(* PLC project GeneratedProgram, SafePLC-Gen SafePLC-Gen Multimodal 1.0 *)
(* stored: creationDateTime 2026-04-25T11:55:04.001507Z *)

PROGRAM GeneratedProgram
  VAR
    FirstScan : BOOL;
    TICSA_4750_03_Scaled : REAL;
    PICSA_4712_02_Scaled : REAL;
    PI_4712_01_Scaled : REAL;
    TICSA_4750_03_EU_Min : REAL;
    TICSA_4750_03_EU_Span : REAL;
    PICSA_4712_02_EU_Min : REAL;
    PICSA_4712_02_EU_Span : REAL;
    PI_4712_01_EU_Min : REAL;
    PI_4712_01_EU_Span : REAL;
    TICSA_4750_03_HH_SP : REAL;
    TICSA_4750_03_H_SP : REAL;
    TICSA_4750_03_L_SP : REAL;
    TICSA_4750_03_LL_SP : REAL;
    TICSA_4750_03_Deadband : REAL;
    PICSA_4712_02_HH_SP : REAL;
    PICSA_4712_02_H_SP : REAL;
    PICSA_4712_02_L_SP : REAL;
    PICSA_4712_02_LL_SP : REAL;
    PICSA_4712_02_Deadband : REAL;
    PI_4712_01_HH_SP : REAL;
    PI_4712_01_H_SP : REAL;
    PI_4712_01_L_SP : REAL;
    PI_4712_01_LL_SP : REAL;
    PI_4712_01_Deadband : REAL;
    TICSA_4750_03_HH_Ack : BOOL;
    TICSA_4750_03_LL_Ack : BOOL;
    PICSA_4712_02_HH_Ack : BOOL;
    PICSA_4712_02_LL_Ack : BOOL;
    PI_4712_01_HH_Ack : BOOL;
    PI_4712_01_LL_Ack : BOOL;
    TICSA_4750_03_LL_Latched : BOOL;
    PICSA_4712_02_HH_Latched : BOOL;
    PICSA_4712_02_LL_Latched : BOOL;
    PI_4712_01_HH_Latched : BOOL;
    PI_4712_01_LL_Latched : BOOL;
    TICSA_4750_03_HH : BOOL;
    TICSA_4750_03_LL : BOOL;
    TICSA_4750_03_H : BOOL;
    TICSA_4750_03_L : BOOL;
    PICSA_4712_02_HH : BOOL;
    PICSA_4712_02_LL : BOOL;
    PICSA_4712_02_H : BOOL;
    PICSA_4712_02_L : BOOL;
    PI_4712_01_HH : BOOL;
    PI_4712_01_LL : BOOL;
    PI_4712_01_H : BOOL;
    PI_4712_01_L : BOOL;
    LOOP_4750_03_TRIP : BOOL;
    LOOP_4712_02_TRIP : BOOL;
    LOOP_104_01_TRIP : BOOL;
    SV_104_01_HH : BOOL;
    SV_104_01_LL : BOOL;
    SAFE_STATE : BOOL;
    TIC_SP : REAL;
    TIC_Error : REAL;
    TIC_Integral : REAL;
    TIC_Kp : REAL;
    TIC_Ki : REAL;
    TIC_Output : REAL;
    PIC_SP : REAL;
    PIC_Error : REAL;
    PIC_Integral : REAL;
    PIC_Kp : REAL;
    PIC_Ki : REAL;
    PIC_Output : REAL;
    HV_MNb_47121 : BOOL;
    HV_MNb_47122 : BOOL;
    HV_75SA21 : BOOL;
    CV_73KH12_50_inlet : BOOL;
    HV_MNc_47125_block : BOOL;
    HV_MNc_47126 : BOOL;
    HV_73KH12_50_main : BOOL;
    HV_QSa_47140 : BOOL;
    HV_QSb_47141 : BOOL;
    HV_MNc_47127_Q80 : BOOL;
    HV_66KL21 : BOOL;
    HV_73KH12_25_PI : BOOL;
    HV_73KH12_25_PICSA : BOOL;
    SV_104_01_Out : BOOL;
    System_Alarm : BOOL;
  END_VAR

            IF FirstScan THEN
    LOOP_4750_03_TRIP    := TRUE;
    LOOP_4712_02_TRIP    := TRUE;
    LOOP_104_01_TRIP     := TRUE;
    SAFE_STATE           := TRUE;
    TV_4750_03_Out       := 6554;
    PV_4712_02_Out       := 6554;
    XV_4750_01           := FALSE;
    SV_104_01_Out        := FALSE;
    HV_MNb_47121         := FALSE;
    HV_MNb_47122         := FALSE;
    HV_75SA21            := FALSE;
    CV_73KH12_50_inlet   := FALSE;
    HV_MNc_47125_block   := FALSE;
    HV_MNc_47126         := FALSE;
    HV_73KH12_50_main    := FALSE;
    HV_QSa_47140         := FALSE;
    HV_QSb_47141         := FALSE;
    HV_MNc_47127_Q80     := FALSE;
    HV_66KL21            := FALSE;
    HV_73KH12_25_PI      := FALSE;
    HV_73KH12_25_PICSA   := FALSE;
    TIC_Integral         := 50.0;
    PIC_Integral         := 50.0;
    TICSA_4750_03_HH_Latched := FALSE;
    TICSA_4750_03_LL_Latched := FALSE;
    PICSA_4712_02_HH_Latched := FALSE;
    PICSA_4712_02_LL_Latched := FALSE;
    PI_4712_01_HH_Latched    := FALSE;
    PI_4712_01_LL_Latched    := FALSE;
    FirstScan            := FALSE;
    RETURN;
END_IF;

TICSA_4750_03_Scaled := ((INT_TO_REAL(TICSA_4750_03_Raw) - 6554.0) / (32767.0 - 6554.0)) * TICSA_4750_03_EU_Span + TICSA_4750_03_EU_Min;
PICSA_4712_02_Scaled := ((INT_TO_REAL(PICSA_4712_02_Raw) - 6554.0) / (32767.0 - 6554.0)) * PICSA_4712_02_EU_Span + PICSA_4712_02_EU_Min;
PI_4712_01_Scaled    := ((INT_TO_REAL(PI_4712_01_Raw)    - 6554.0) / (32767.0 - 6554.0)) * PI_4712_01_EU_Span    + PI_4712_01_EU_Min;

(* TICSA-4750.03 HH latching alarm *)
IF TICSA_4750_03_Scaled >= TICSA_4750_03_HH_SP THEN
    TICSA_4750_03_HH_Latched := TRUE;
ELSIF TICSA_4750_03_HH_Ack AND (TICSA_4750_03_Scaled <= (TICSA_4750_03_HH_SP - TICSA_4750_03_Deadband)) THEN
    TICSA_4750_03_HH_Latched := FALSE;
END_IF;
TICSA_4750_03_HH := TICSA_4750_03_HH_Latched;

(* TICSA-4750.03 LL latching alarm *)
IF TICSA_4750_03_Scaled <= TICSA_4750_03_LL_SP THEN
    TICSA_4750_03_LL_Latched := TRUE;
ELSIF TICSA_4750_03_LL_Ack AND (TICSA_4750_03_Scaled >= (TICSA_4750_03_LL_SP + TICSA_4750_03_Deadband)) THEN
    TICSA_4750_03_LL_Latched := FALSE;
END_IF;
TICSA_4750_03_LL := TICSA_4750_03_LL_Latched;

(* TICSA-4750.03 H/L non-latching *)
IF TICSA_4750_03_Scaled >= TICSA_4750_03_H_SP THEN
    TICSA_4750_03_H := TRUE;
ELSIF TICSA_4750_03_Scaled <= (TICSA_4750_03_H_SP - TICSA_4750_03_Deadband) THEN
    TICSA_4750_03_H := FALSE;
END_IF;

IF TICSA_4750_03_Scaled <= TICSA_4750_03_L_SP THEN
    TICSA_4750_03_L := TRUE;
ELSIF TICSA_4750_03_Scaled >= (TICSA_4750_03_L_SP + TICSA_4750_03_Deadband) THEN
    TICSA_4750_03_L := FALSE;
END_IF;

(* PICSA-4712.02 HH latching alarm *)
IF PICSA_4712_02_Scaled >= PICSA_4712_02_HH_SP THEN
    PICSA_4712_02_HH_Latched := TRUE;
ELSIF PICSA_4712_02_HH_Ack AND (PICSA_4712_02_Scaled <= (PICSA_4712_02_HH_SP - PICSA_4712_02_Deadband)) THEN
    PICSA_4712_02_HH_Latched := FALSE;
END_IF;
PICSA_4712_02_HH := PICSA_4712_02_HH_Latched;

(* PICSA-4712.02 LL latching alarm *)
IF PICSA_4712_02_Scaled <= PICSA_4712_02_LL_SP THEN
    PICSA_4712_02_LL_Latched := TRUE;
ELSIF PICSA_4712_02_LL_Ack AND (PICSA_4712_02_Scaled >= (PICSA_4712_02_LL_SP + PICSA_4712_02_Deadband)) THEN
    PICSA_4712_02_LL_Latched := FALSE;
END_IF;
PICSA_4712_02_LL := PICSA_4712_02_LL_Latched;

(* PICSA-4712.02 H/L non-latching *)
IF PICSA_4712_02_Scaled >= PICSA_4712_02_H_SP THEN
    PICSA_4712_02_H := TRUE;
ELSIF PICSA_4712_02_Scaled <= (PICSA_4712_02_H_SP - PICSA_4712_02_Deadband) THEN
    PICSA_4712_02_H := FALSE;
END_IF;

IF PICSA_4712_02_Scaled <= PICSA_4712_02_L_SP THEN
    PICSA_4712_02_L := TRUE;
ELSIF PICSA_4712_02_Scaled >= (PICSA_4712_02_L_SP + PICSA_4712_02_Deadband) THEN
    PICSA_4712_02_L := FALSE;
END_IF;

(* PI-4712.01 HH latching alarm *)
IF PI_4712_01_Scaled >= PI_4712_01_HH_SP THEN
    PI_4712_01_HH_Latched := TRUE;
ELSIF PI_4712_01_HH_Ack AND (PI_4712_01_Scaled <= (PI_4712_01_HH_SP - PI_4712_01_Deadband)) THEN
    PI_4712_01_HH_Latched := FALSE;
END_IF;
PI_4712_01_HH := PI_4712_01_HH_Latched;

(* PI-4712.01 LL latching alarm *)
IF PI_4712_01_Scaled <= PI_4712_01_LL_SP THEN
    PI_4712_01_LL_Latched := TRUE;
ELSIF PI_4712_01_LL_Ack AND (PI_4712_01_Scaled >= (PI_4712_01_LL_SP + PI_4712_01_Deadband)) THEN
    PI_4712_01_LL_Latched := FALSE;
END_IF;
PI_4712_01_LL := PI_4712_01_LL_Latched;

(* PI-4712.01 H/L non-latching *)
IF PI_4712_01_Scaled >= PI_4712_01_H_SP THEN
    PI_4712_01_H := TRUE;
ELSIF PI_4712_01_Scaled <= (PI_4712_01_H_SP - PI_4712_01_Deadband) THEN
    PI_4712_01_H := FALSE;
END_IF;

IF PI_4712_01_Scaled <= PI_4712_01_L_SP THEN
    PI_4712_01_L := TRUE;
ELSIF PI_4712_01_Scaled >= (PI_4712_01_L_SP + PI_4712_01_Deadband) THEN
    PI_4712_01_L := FALSE;
END_IF;

(* Safety trip latches *)
IF TICSA_4750_03_HH OR TICSA_4750_03_LL THEN
    LOOP_4750_03_TRIP := TRUE;
ELSIF LOOP_4750_03_TRIP AND MANUAL_RESET AND NOT TICSA_4750_03_HH AND NOT TICSA_4750_03_LL THEN
    LOOP_4750_03_TRIP := FALSE;
END_IF;

IF PICSA_4712_02_HH OR PICSA_4712_02_LL THEN
    LOOP_4712_02_TRIP := TRUE;
ELSIF LOOP_4712_02_TRIP AND MANUAL_RESET AND NOT PICSA_4712_02_HH AND NOT PICSA_4712_02_LL THEN
    LOOP_4712_02_TRIP := FALSE;
END_IF;

IF SV_104_01_HH OR SV_104_01_LL THEN
    LOOP_104_01_TRIP := TRUE;
ELSIF LOOP_104_01_TRIP AND MANUAL_RESET AND NOT SV_104_01_HH AND NOT SV_104_01_LL THEN
    LOOP_104_01_TRIP := FALSE;
END_IF;

SAFE_STATE := ESTOP OR LOOP_4750_03_TRIP OR LOOP_4712_02_TRIP OR LOOP_104_01_TRIP;

IF NOT SAFE_STATE THEN
    TIC_Error    := TIC_SP - TICSA_4750_03_Scaled;
    TIC_Integral := TIC_Integral + (TIC_Ki * TIC_Error);
    IF TIC_Integral > 100.0 THEN
        TIC_Integral := 100.0;
    ELSIF TIC_Integral < 0.0 THEN
        TIC_Integral := 0.0;
    END_IF;
    TIC_Output := (TIC_Kp * TIC_Error) + TIC_Integral;
    IF TIC_Output > 100.0 THEN
        TIC_Output := 100.0;
    ELSIF TIC_Output < 0.0 THEN
        TIC_Output := 0.0;
    END_IF;
    TV_4750_03_Out := REAL_TO_INT(6554.0 + (TIC_Output / 100.0) * (32767.0 - 6554.0));

    PIC_Error    := PIC_SP - PICSA_4712_02_Scaled;
    PIC_Integral := PIC_Integral + (PIC_Ki * PIC_Error);
    IF PIC_Integral > 100.0 THEN
        PIC_Integral := 100.0;
    ELSIF PIC_Integral < 0.0 THEN
        PIC_Integral := 0.0;
    END_IF;
    PIC_Output := (PIC_Kp * PIC_Error) + PIC_Integral;
    IF PIC_Output > 100.0 THEN
        PIC_Output := 100.0;
    ELSIF PIC_Output < 0.0 THEN
        PIC_Output := 0.0;
    END_IF;
    PV_4712_02_Out := REAL_TO_INT(6554.0 + (PIC_Output / 100.0) * (32767.0 - 6554.0));

    XV_4750_01         := HS_4750_01;
    SV_104_01_Out      := TRUE;
    HV_MNb_47121       := TRUE;
    HV_MNb_47122       := TRUE;
    HV_75SA21          := TRUE;
    CV_73KH12_50_inlet := TRUE;
    HV_MNc_47125_block := TRUE;
    HV_MNc_47126       := TRUE;
    HV_73KH12_50_main  := TRUE;
    HV_QSa_47140       := TRUE;
    HV_QSb_47141       := TRUE;
    HV_MNc_47127_Q80   := TRUE;
    HV_66KL21          := TRUE;
    HV_73KH12_25_PI    := TRUE;
    HV_73KH12_25_PICSA := TRUE;
ELSE
    TV_4750_03_Out     := 6554;
    PV_4712_02_Out     := 6554;
    XV_4750_01         := FALSE;
    SV_104_01_Out      := FALSE;
    HV_MNb_47121       := FALSE;
    HV_MNb_47122       := FALSE;
    HV_75SA21          := FALSE;
    CV_73KH12_50_inlet := FALSE;
    HV_MNc_47125_block := FALSE;
    HV_MNc_47126       := FALSE;
    HV_73KH12_50_main  := FALSE;
    HV_QSa_47140       := FALSE;
    HV_QSb_47141       := FALSE;
    HV_MNc_47127_Q80   := FALSE;
    HV_66KL21          := FALSE;
    HV_73KH12_25_PI    := FALSE;
    HV_73KH12_25_PICSA := FALSE;
END_IF;

System_Alarm :=
    TICSA_4750_03_HH_Latched OR TICSA_4750_03_LL_Latched OR
    TICSA_4750_03_H          OR TICSA_4750_03_L          OR
    PICSA_4712_02_HH_Latched OR PICSA_4712_02_LL_Latched OR
    PICSA_4712_02_H          OR PICSA_4712_02_L          OR
    PI_4712_01_HH_Latched    OR PI_4712_01_LL_Latched    OR
    PI_4712_01_H             OR PI_4712_01_L             OR
    LOOP_4750_03_TRIP        OR LOOP_4712_02_TRIP        OR
    LOOP_104_01_TRIP         OR SAFE_STATE;
          
END_PROGRAM

CONFIGURATION Config0
  RESOURCE Res0 ON PLC
    TASK MainTask(INTERVAL := T#20ms, PRIORITY := 0);
    PROGRAM Main : GeneratedProgram;
  END_RESOURCE
END_CONFIGURATION
